(* Logix 5000 project; controller _1407974_PSG_7315 vendor 1 type 14 code 154 rev 20.11; software revision 20.06; part 3 of 4 *)
(* tags used below, declared in another part *)
   AI_L_2_0_Pure_Steam_Conductivity : Analog_Input;
   AI_L_2_1_FW_Press_Low_Warning : OIT_Set_Point_Entry;
   AI_L_2_1_FW_Pressure : Analog_Input;
   AI_R_2_0_Pure_Steam_Temperature : Analog_Input;
   AI_R_2_1_Cond_Pure_Steam_Temperature : Analog_Input;
   Alarm_Pure_Steam_High_Temperature : ALIAS FOR Alarms_Warnings.Latch_Bit[0].4;
   Alarm_Pure_Steam_Temp_Error_Timer : TIMER;
   Alarm_Pure_Steam_Temp_Input_Error : ALIAS FOR Alarms_Warnings.Latch_Bit[0].5;
   Alarm_Pure_Steam_Temp_Input_Error_Ack : ALIAS FOR Alarms_Warnings.Ack[0].5;
   Alarm_Separator_High_Level : ALIAS FOR Alarms_Warnings.Latch_Bit[0].2;
   Alarm_Separator_Low_Level : ALIAS FOR Alarms_Warnings.Latch_Bit[0].3;
   Alarms_Warnings : AW;
   AO_L_3_0_VFD_SPEED : Analog_Output;
   AO_L_3_1_Available : Analog_Output;
   AO_L_3_2_Available : Analog_Output;
   AO_L_3_3_Available : Analog_Output;
   AO_R_4_0_Pure_Steam_Temperature : Analog_Output;
   AO_R_4_1_Available : Analog_Output;
   Cond_Pure_Steam_Hi_Cond_Set_Point_Entry : OIT_Set_Point_Entry;
   Cond_Pure_Steam_Hi_Temp_Set_Point_Entry : OIT_Set_Point_Entry;
   DI_R_1_0_Hi_Hi_Level_LSHH_1950 : ALIAS FOR DI_Remote_1.0;
   DI_R_1_3_Low_Level_LSL_1950 : ALIAS FOR DI_Remote_1.3;
   DI_R_1_4_Air_Low_Pressure_PSL_4030 : ALIAS FOR DI_Remote_1.4;
   DO_L_1_14_Feed_Water_Pump_Contactor : Discrete_Out;
   DO_L_1_1_Alarm_Horn : Discrete_Out;
   DO_L_1_2_Alarm_Light : Discrete_Out;
   DO_Local_1 : INT;
   Feed_Water_Pressure_Set_Point_Entry : OIT_Set_Point_Entry;
   Feedwater_Pressure_PID : PID;
   Free_Run_Pulse_Timer : TIMER;
   FW_Press_PID_Gain_Set_Point_Entry : OIT_Set_Point_Entry;
   FW_Press_PID_Manual_Output_Entry : OIT_Set_Point_Entry;
   FW_Press_PID_Rate_Set_Point_Entry : OIT_Set_Point_Entry;
   FW_Press_PID_Reset_SetPoint_Entry : OIT_Set_Point_Entry;
   FW_Press_PID_Temp_Set_Point_Entry : OIT_Set_Point_Entry;
   Lamp_Test : Push_Button;
   Local_Remote : Latched_Push_Button;
   Low_Feedwater_Pressure : BOOL;
   Network_Ack_All : BOOL;
   Network_Silence : BOOL;
   OIT : OIT_Connections;
   OIT_Auto_Time_Date_Sync : TIMER;
   OIT_Auto_Time_Date_Sync_Interval : TIMER;
   OIT_Day_Set : Push_Button;
   OIT_Hour_Set : Push_Button;
   OIT_Message : OIT_Message;
   OIT_Minute_Set : Push_Button;
   OIT_Month_Set : Push_Button;
   OIT_Year_Set : Push_Button;
   PID_Ramp_Time_Seconds : DINT;
   PID_Ramp_Timer : TIMER;
   Pulse_Bit : BOOL;
   Pure_Steam_High_Temp_Set_Point_Entry : OIT_Set_Point_Entry;
   Pure_Steam_Low_Temp_Set_Point_Entry : OIT_Set_Point_Entry;
   Pure_Steam_Temp_PID_Gain_Set_Point_Entry : OIT_Set_Point_Entry;
   Pure_Steam_Temp_PID_Manual_Output_Entry : OIT_Set_Point_Entry;
   Pure_Steam_Temp_PID_Ramp_Time_Entry : OIT_Set_Point_Entry;
   Pure_Steam_Temp_PID_Rate_Set_Point_Entry : OIT_Set_Point_Entry;
   Pure_Steam_Temp_PID_Reset_SetPoint_Entry : OIT_Set_Point_Entry;
   Pure_Steam_Temp_PID_Temp_Set_Point_Entry : OIT_Set_Point_Entry;
   Pure_Steam_Temperature : PID;
   Pure_Steam_Temperature_Set_Point_Entry : OIT_Set_Point_Entry;
   Read_PLC_Clock : DINT[7];
   Set_PLC_Clock : DINT[7];
   Unit_Hot : BOOL;
   Unit_Status : Unit_Status;
   VFD_Relay_Input : BOOL;
   Warning_Air_Low_Pressure_Timer : TIMER;
   Warning_Cond_Pure_Steam_Analyzer_Fault : ALIAS FOR Alarms_Warnings.Latch_Bit[1].4;
   Warning_Cond_Pure_Steam_Conductivity : ALIAS FOR Alarms_Warnings.Latch_Bit[1].3;
   Warning_Feedwater_Low_Pressure : ALIAS FOR Alarms_Warnings.Latch_Bit[1].9;
   Warning_Feedwater_Press_Low_Pressure_Ack : ALIAS FOR Alarms_Warnings.Ack[1].9;
   Warning_FW_Press_Low_Pressure_Timer : TIMER;
   Warning_Instrument_Air_Low_Pressure : ALIAS FOR Alarms_Warnings.Latch_Bit[1].2;
   Warning_Instrument_Air_Low_Pressure_Ack : ALIAS FOR Alarms_Warnings.Ack[1].2;
   Warning_PLC_OIT_Comm_Counter : COUNTER;
   Warning_PLC_OIT_Comm_Timer : TIMER;
   Warning_PLC_OIT_Commuications_Ack : ALIAS FOR Alarms_Warnings.Ack[1].0;
   Warning_PLC_OIT_Communications : ALIAS FOR Alarms_Warnings.Latch_Bit[1].0;
   Warning_Pure_Steam_Low_Temp_Timer_A : TIMER;
   Warning_Pure_Steam_Low_Temp_Timer_B : TIMER;
   Warning_Pure_Steam_Low_Temperature : ALIAS FOR Alarms_Warnings.Latch_Bit[1].7;
   Warning_Pure_Steam_Low_Temperature_Ack : ALIAS FOR Alarms_Warnings.Ack[1].7;
(* MainProgram, continued *)

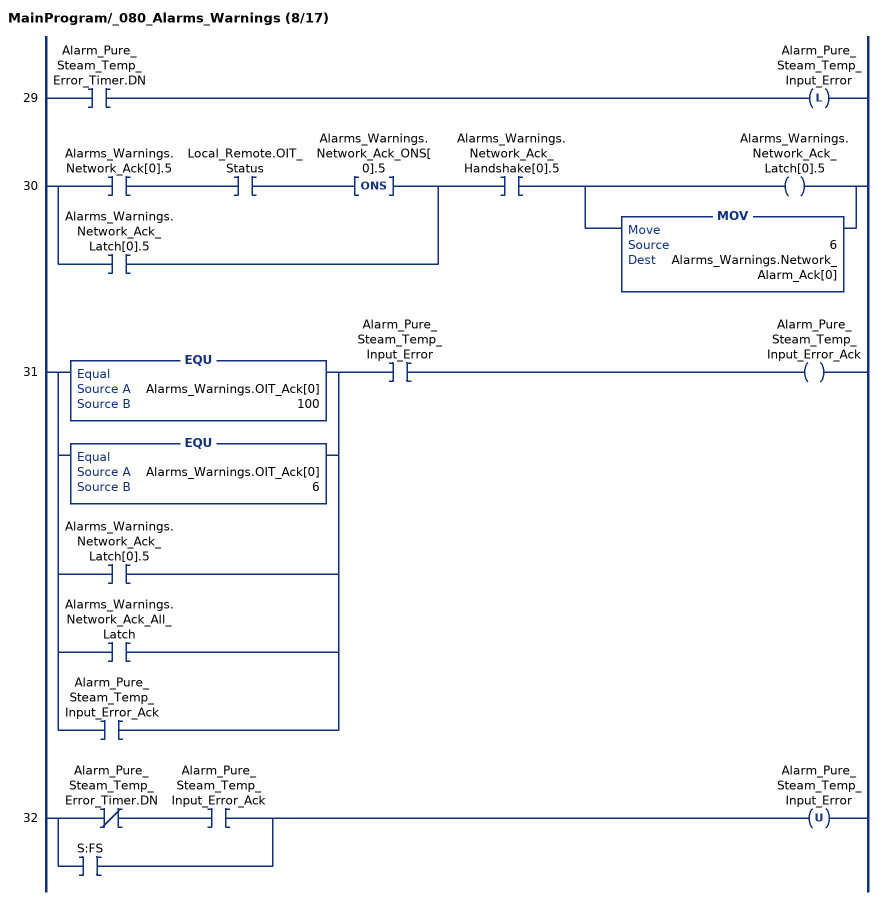
   [picture p43: MainProgram/_080_Alarms_Warnings rungs 29-32]
   29: XIC(Alarm_Pure_Steam_Temp_Error_Timer.DN)OTL(Alarm_Pure_Steam_Temp_Input_Error);
   30: [XIC(Alarms_Warnings.Network_Ack[0].5) XIC(Local_Remote.OIT_Status) ONS(Alarms_Warnings.Network_Ack_ONS[0].5) ,XIC(Alarms_Warnings.Network_Ack_Latch[0].5) ]XIC(Alarms_Warnings.Network_Ack_Handshake[0].5)[OTE(Alarms_Warnings.Network_Ack_Latch[0].5) ,MOV(6,Alarms_Warnings.Network_Alarm_Ack[0]) ];
   31: [EQU(Alarms_Warnings.OIT_Ack[0],100) ,EQU(Alarms_Warnings.OIT_Ack[0],6) ,XIC(Alarms_Warnings.Network_Ack_Latch[0].5) ,XIC(Alarms_Warnings.Network_Ack_All_Latch) ,XIC(Alarm_Pure_Steam_Temp_Input_Error_Ack) ]XIC(Alarm_Pure_Steam_Temp_Input_Error)OTE(Alarm_Pure_Steam_Temp_Input_Error_Ack);
   32: [XIO(Alarm_Pure_Steam_Temp_Error_Timer.DN) XIC(Alarm_Pure_Steam_Temp_Input_Error_Ack) ,XIC(S:FS) ]OTU(Alarm_Pure_Steam_Temp_Input_Error);
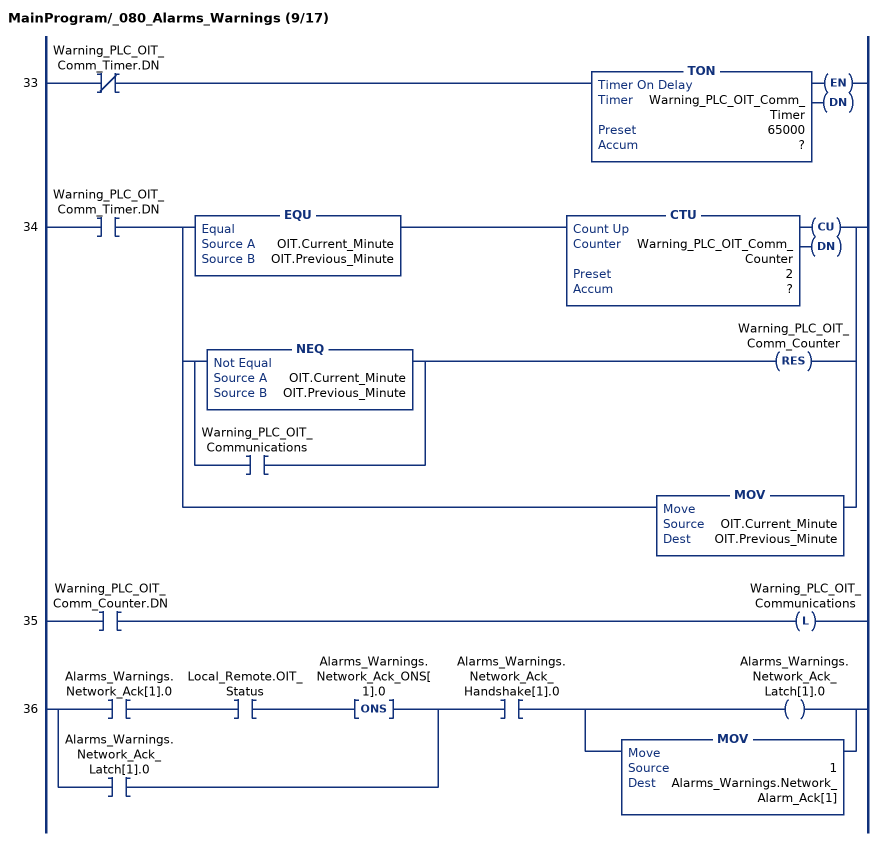
   33: XIO(Warning_PLC_OIT_Comm_Timer.DN)TON(Warning_PLC_OIT_Comm_Timer,?,?);
   34: XIC(Warning_PLC_OIT_Comm_Timer.DN)[EQU(OIT.Current_Minute,OIT.Previous_Minute) CTU(Warning_PLC_OIT_Comm_Counter,?,?) ,[NEQ(OIT.Current_Minute,OIT.Previous_Minute) ,XIC(Warning_PLC_OIT_Communications) ] RES(Warning_PLC_OIT_Comm_Counter) ,MOV(OIT.Current_Minute,OIT.Previous_Minute) ];
   35: XIC(Warning_PLC_OIT_Comm_Counter.DN)OTL(Warning_PLC_OIT_Communications);
   36: [XIC(Alarms_Warnings.Network_Ack[1].0) XIC(Local_Remote.OIT_Status) ONS(Alarms_Warnings.Network_Ack_ONS[1].0) ,XIC(Alarms_Warnings.Network_Ack_Latch[1].0) ]XIC(Alarms_Warnings.Network_Ack_Handshake[1].0)[OTE(Alarms_Warnings.Network_Ack_Latch[1].0) ,MOV(1,Alarms_Warnings.Network_Alarm_Ack[1]) ];
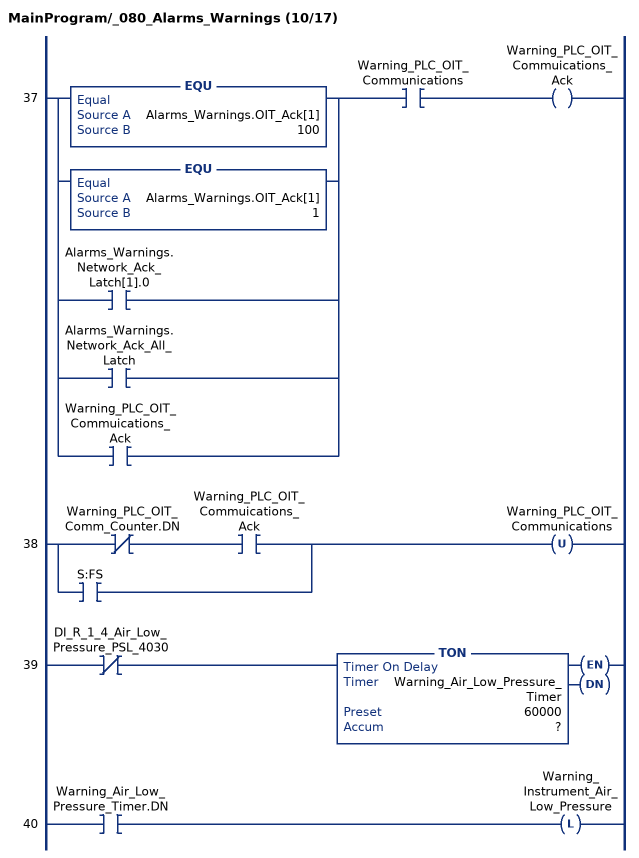
   37: [EQU(Alarms_Warnings.OIT_Ack[1],100) ,EQU(Alarms_Warnings.OIT_Ack[1],1) ,XIC(Alarms_Warnings.Network_Ack_Latch[1].0) ,XIC(Alarms_Warnings.Network_Ack_All_Latch) ,XIC(Warning_PLC_OIT_Commuications_Ack) ]XIC(Warning_PLC_OIT_Communications)OTE(Warning_PLC_OIT_Commuications_Ack);
   38: [XIO(Warning_PLC_OIT_Comm_Counter.DN) XIC(Warning_PLC_OIT_Commuications_Ack) ,XIC(S:FS) ]OTU(Warning_PLC_OIT_Communications);
   39: XIO(DI_R_1_4_Air_Low_Pressure_PSL_4030)TON(Warning_Air_Low_Pressure_Timer,?,?);
   40: XIC(Warning_Air_Low_Pressure_Timer.DN)OTL(Warning_Instrument_Air_Low_Pressure);
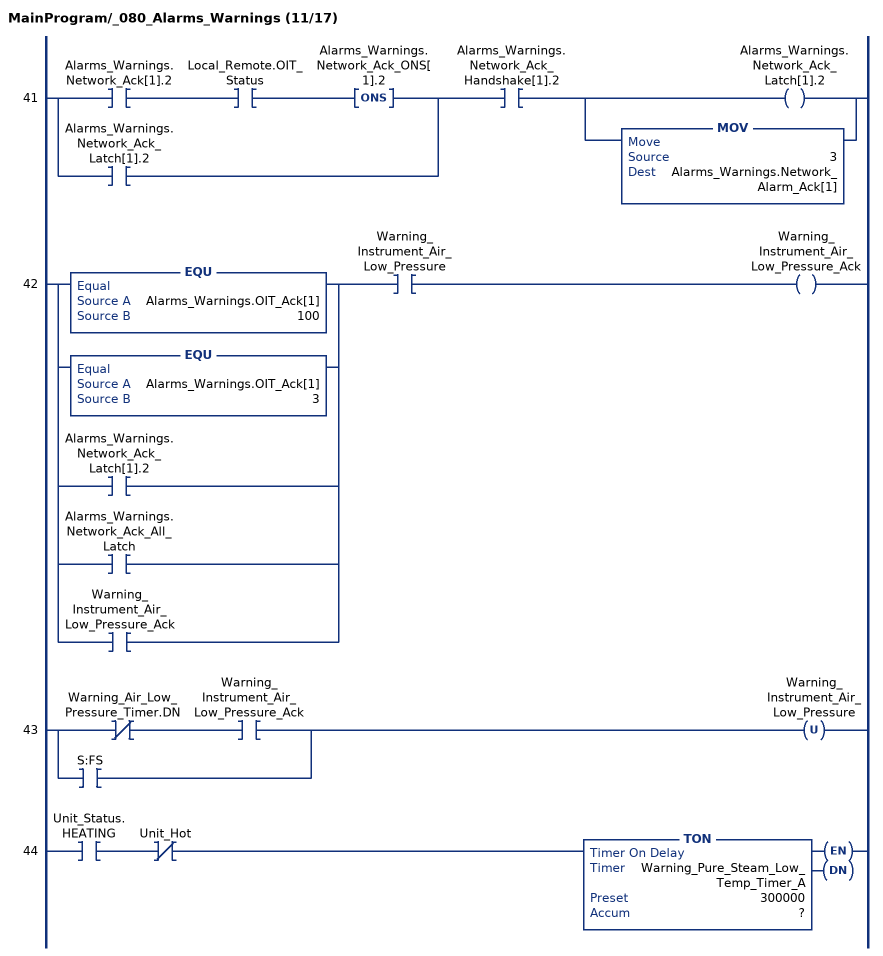
   41: [XIC(Alarms_Warnings.Network_Ack[1].2) XIC(Local_Remote.OIT_Status) ONS(Alarms_Warnings.Network_Ack_ONS[1].2) ,XIC(Alarms_Warnings.Network_Ack_Latch[1].2) ]XIC(Alarms_Warnings.Network_Ack_Handshake[1].2)[OTE(Alarms_Warnings.Network_Ack_Latch[1].2) ,MOV(3,Alarms_Warnings.Network_Alarm_Ack[1]) ];
   42: [EQU(Alarms_Warnings.OIT_Ack[1],100) ,EQU(Alarms_Warnings.OIT_Ack[1],3) ,XIC(Alarms_Warnings.Network_Ack_Latch[1].2) ,XIC(Alarms_Warnings.Network_Ack_All_Latch) ,XIC(Warning_Instrument_Air_Low_Pressure_Ack) ]XIC(Warning_Instrument_Air_Low_Pressure)OTE(Warning_Instrument_Air_Low_Pressure_Ack);
   43: [XIO(Warning_Air_Low_Pressure_Timer.DN) XIC(Warning_Instrument_Air_Low_Pressure_Ack) ,XIC(S:FS) ]OTU(Warning_Instrument_Air_Low_Pressure);
   44: XIC(Unit_Status.HEATING)XIO(Unit_Hot)TON(Warning_Pure_Steam_Low_Temp_Timer_A,?,?);
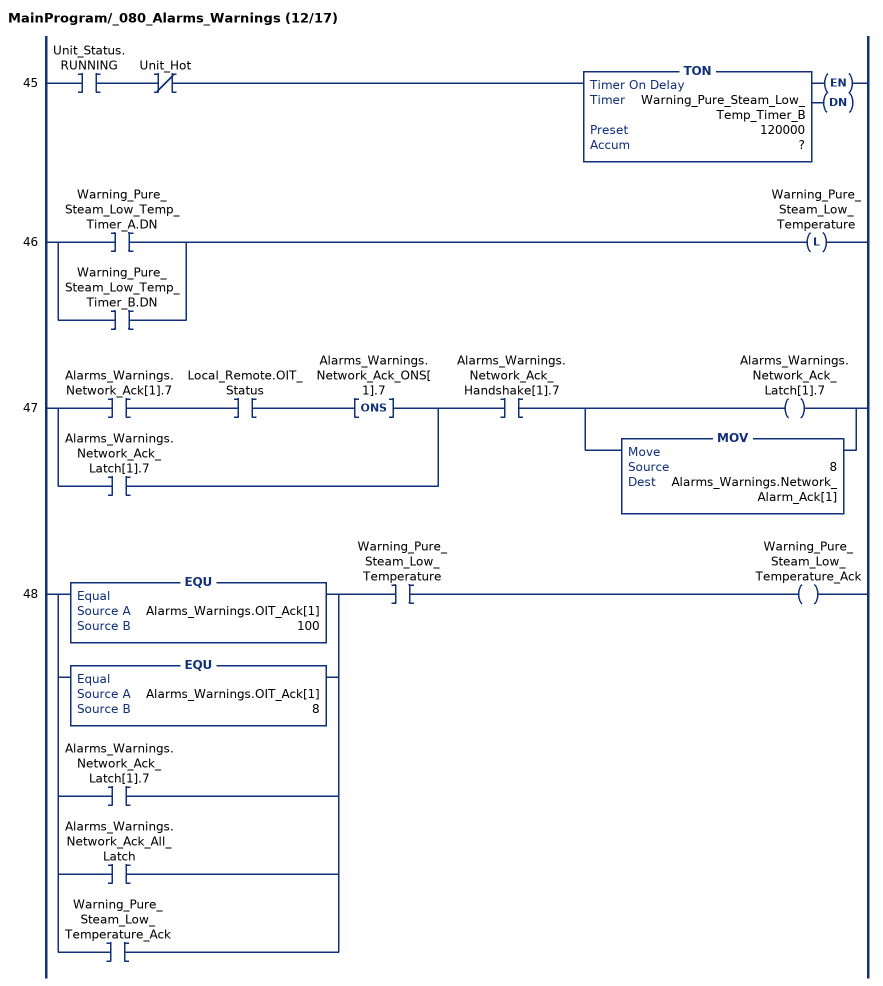
   45: XIC(Unit_Status.RUNNING)XIO(Unit_Hot)TON(Warning_Pure_Steam_Low_Temp_Timer_B,?,?);
   46: [XIC(Warning_Pure_Steam_Low_Temp_Timer_A.DN) ,XIC(Warning_Pure_Steam_Low_Temp_Timer_B.DN) ]OTL(Warning_Pure_Steam_Low_Temperature);
   47: [XIC(Alarms_Warnings.Network_Ack[1].7) XIC(Local_Remote.OIT_Status) ONS(Alarms_Warnings.Network_Ack_ONS[1].7) ,XIC(Alarms_Warnings.Network_Ack_Latch[1].7) ]XIC(Alarms_Warnings.Network_Ack_Handshake[1].7)[OTE(Alarms_Warnings.Network_Ack_Latch[1].7) ,MOV(8,Alarms_Warnings.Network_Alarm_Ack[1]) ];
   48: [EQU(Alarms_Warnings.OIT_Ack[1],100) ,EQU(Alarms_Warnings.OIT_Ack[1],8) ,XIC(Alarms_Warnings.Network_Ack_Latch[1].7) ,XIC(Alarms_Warnings.Network_Ack_All_Latch) ,XIC(Warning_Pure_Steam_Low_Temperature_Ack) ]XIC(Warning_Pure_Steam_Low_Temperature)OTE(Warning_Pure_Steam_Low_Temperature_Ack);
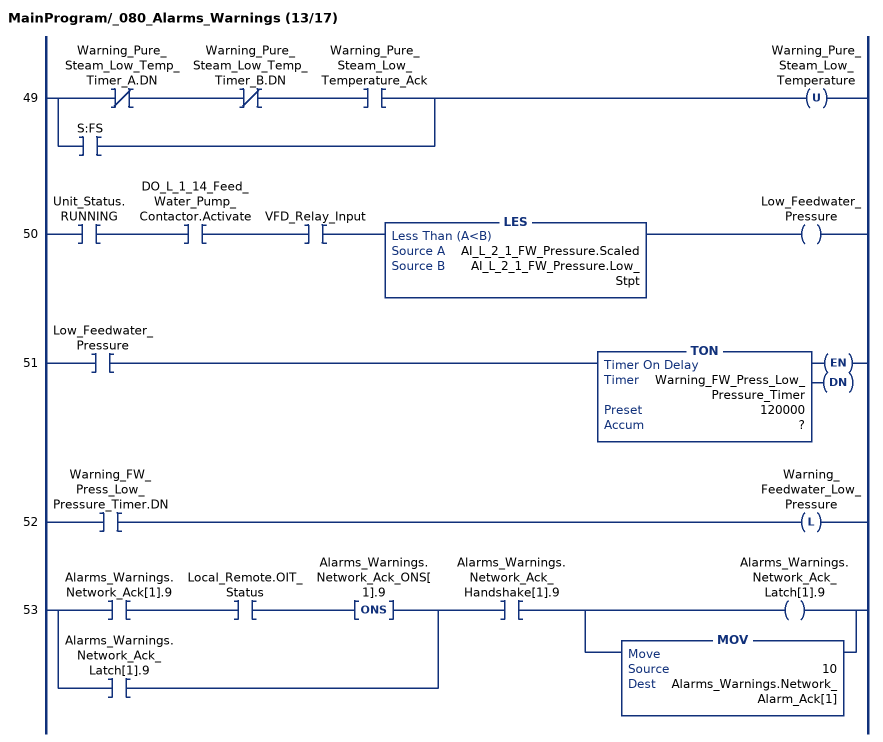
   49: [XIO(Warning_Pure_Steam_Low_Temp_Timer_A.DN) XIO(Warning_Pure_Steam_Low_Temp_Timer_B.DN) XIC(Warning_Pure_Steam_Low_Temperature_Ack) ,XIC(S:FS) ]OTU(Warning_Pure_Steam_Low_Temperature);
   50: XIC(Unit_Status.RUNNING)XIC(DO_L_1_14_Feed_Water_Pump_Contactor.Activate)XIC(VFD_Relay_Input)LES(AI_L_2_1_FW_Pressure.Scaled,AI_L_2_1_FW_Pressure.Low_Stpt)OTE(Low_Feedwater_Pressure);
   51: XIC(Low_Feedwater_Pressure)TON(Warning_FW_Press_Low_Pressure_Timer,?,?);
   52: XIC(Warning_FW_Press_Low_Pressure_Timer.DN)OTL(Warning_Feedwater_Low_Pressure);
   53: [XIC(Alarms_Warnings.Network_Ack[1].9) XIC(Local_Remote.OIT_Status) ONS(Alarms_Warnings.Network_Ack_ONS[1].9) ,XIC(Alarms_Warnings.Network_Ack_Latch[1].9) ]XIC(Alarms_Warnings.Network_Ack_Handshake[1].9)[OTE(Alarms_Warnings.Network_Ack_Latch[1].9) ,MOV(10,Alarms_Warnings.Network_Alarm_Ack[1]) ];
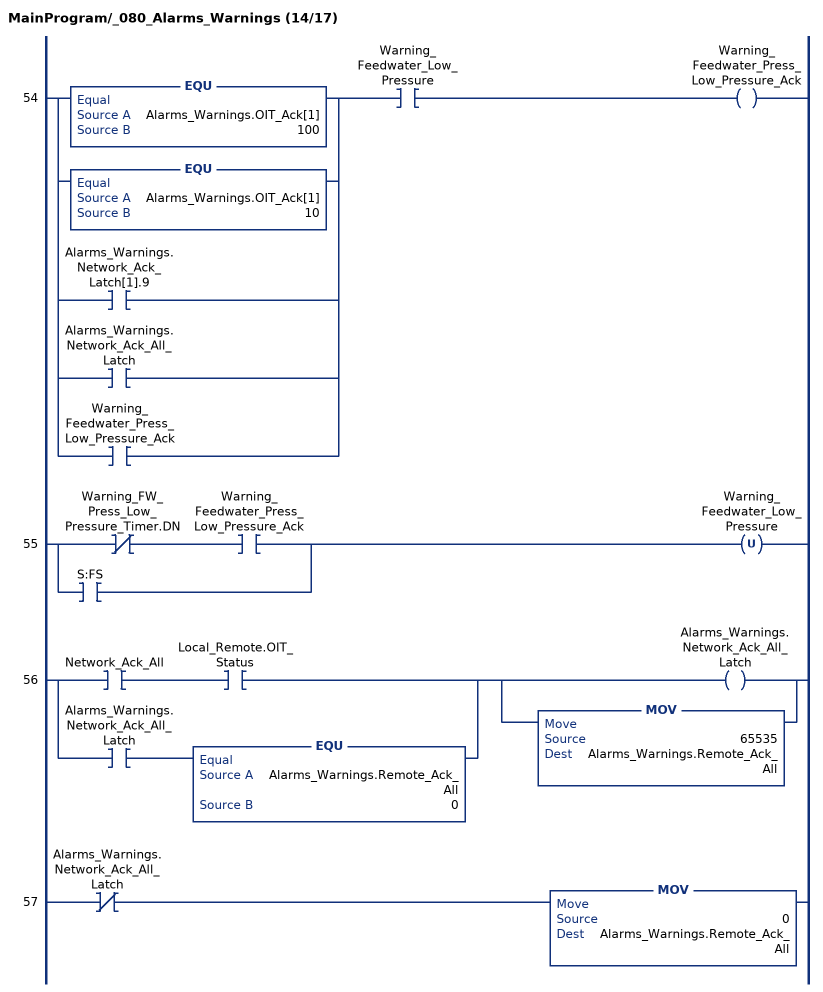
   54: [EQU(Alarms_Warnings.OIT_Ack[1],100) ,EQU(Alarms_Warnings.OIT_Ack[1],10) ,XIC(Alarms_Warnings.Network_Ack_Latch[1].9) ,XIC(Alarms_Warnings.Network_Ack_All_Latch) ,XIC(Warning_Feedwater_Press_Low_Pressure_Ack) ]XIC(Warning_Feedwater_Low_Pressure)OTE(Warning_Feedwater_Press_Low_Pressure_Ack);
   55: [XIO(Warning_FW_Press_Low_Pressure_Timer.DN) XIC(Warning_Feedwater_Press_Low_Pressure_Ack) ,XIC(S:FS) ]OTU(Warning_Feedwater_Low_Pressure);
   56: [XIC(Network_Ack_All) XIC(Local_Remote.OIT_Status) ,XIC(Alarms_Warnings.Network_Ack_All_Latch) EQU(Alarms_Warnings.Remote_Ack_All,0) ][OTE(Alarms_Warnings.Network_Ack_All_Latch) ,MOV(65535,Alarms_Warnings.Remote_Ack_All) ];
   57: XIO(Alarms_Warnings.Network_Ack_All_Latch)MOV(0,Alarms_Warnings.Remote_Ack_All);
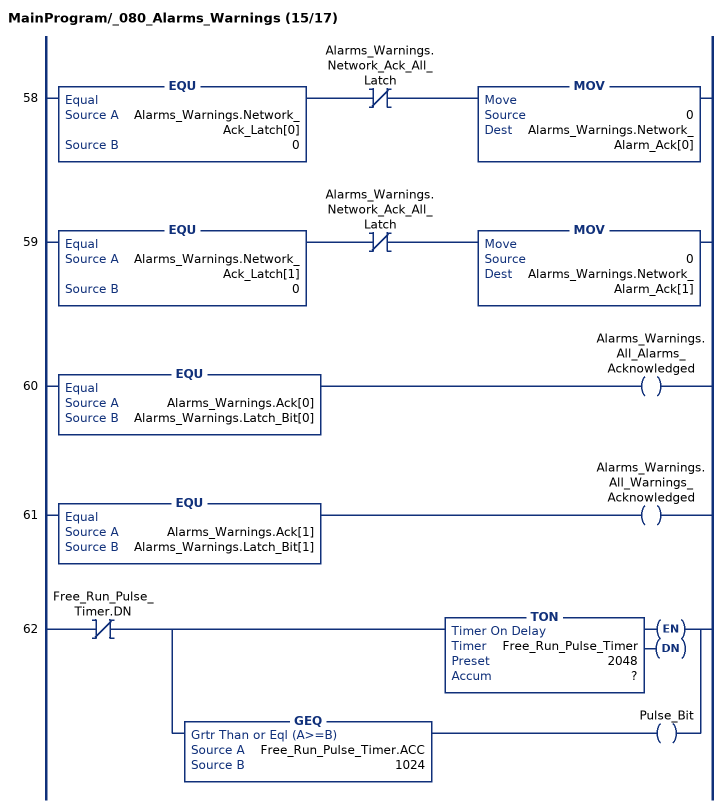
   58: EQU(Alarms_Warnings.Network_Ack_Latch[0],0)XIO(Alarms_Warnings.Network_Ack_All_Latch)MOV(0,Alarms_Warnings.Network_Alarm_Ack[0]);
   59: EQU(Alarms_Warnings.Network_Ack_Latch[1],0)XIO(Alarms_Warnings.Network_Ack_All_Latch)MOV(0,Alarms_Warnings.Network_Alarm_Ack[1]);
   60: EQU(Alarms_Warnings.Ack[0],Alarms_Warnings.Latch_Bit[0])OTE(Alarms_Warnings.All_Alarms_Acknowledged);
   61: EQU(Alarms_Warnings.Ack[1],Alarms_Warnings.Latch_Bit[1])OTE(Alarms_Warnings.All_Warnings_Acknowledged);
   62: XIO(Free_Run_Pulse_Timer.DN)[TON(Free_Run_Pulse_Timer,?,?) ,GEQ(Free_Run_Pulse_Timer.ACC,1024) OTE(Pulse_Bit) ];
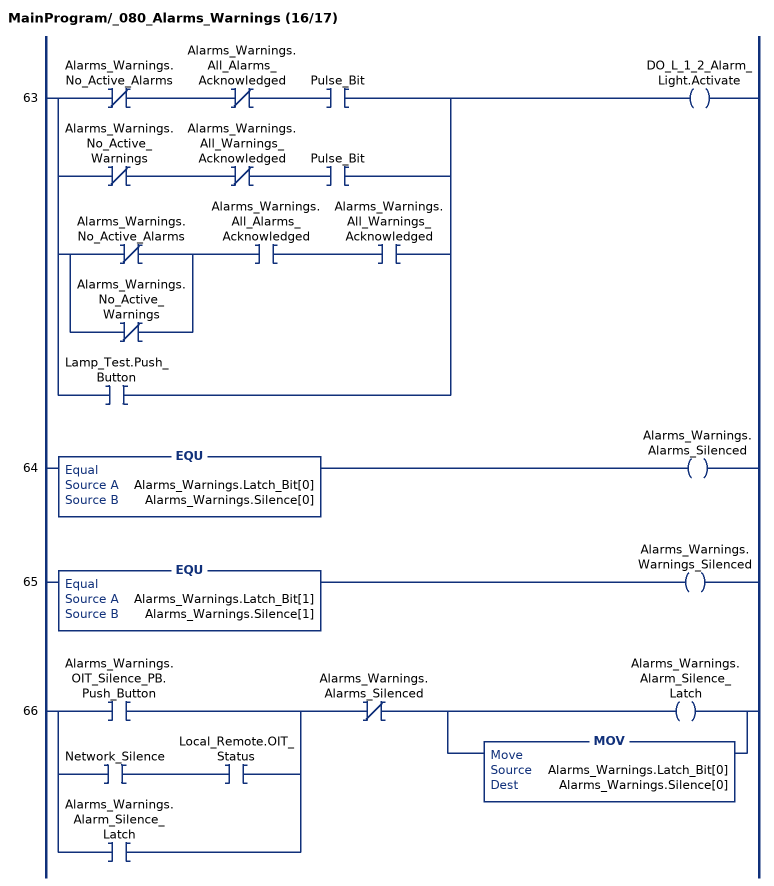
   63: [XIO(Alarms_Warnings.No_Active_Alarms) XIO(Alarms_Warnings.All_Alarms_Acknowledged) XIC(Pulse_Bit) ,XIO(Alarms_Warnings.No_Active_Warnings) XIO(Alarms_Warnings.All_Warnings_Acknowledged) XIC(Pulse_Bit) ,[XIO(Alarms_Warnings.No_Active_Alarms) ,XIO(Alarms_Warnings.No_Active_Warnings) ] XIC(Alarms_Warnings.All_Alarms_Acknowledged) XIC(Alarms_Warnings.All_Warnings_Acknowledged) ,XIC(Lamp_Test.Push_Button) ]OTE(DO_L_1_2_Alarm_Light.Activate);
   64: EQU(Alarms_Warnings.Latch_Bit[0],Alarms_Warnings.Silence[0])OTE(Alarms_Warnings.Alarms_Silenced);
   65: EQU(Alarms_Warnings.Latch_Bit[1],Alarms_Warnings.Silence[1])OTE(Alarms_Warnings.Warnings_Silenced);
   66: [XIC(Alarms_Warnings.OIT_Silence_PB.Push_Button) ,XIC(Network_Silence) XIC(Local_Remote.OIT_Status) ,XIC(Alarms_Warnings.Alarm_Silence_Latch) ]XIO(Alarms_Warnings.Alarms_Silenced)[OTE(Alarms_Warnings.Alarm_Silence_Latch) ,MOV(Alarms_Warnings.Latch_Bit[0],Alarms_Warnings.Silence[0]) ];
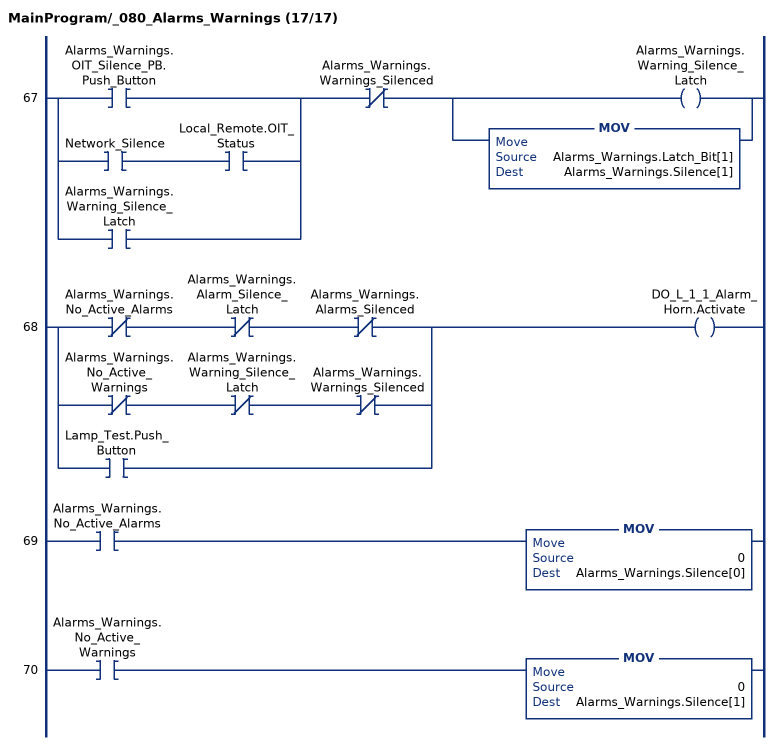
   67: [XIC(Alarms_Warnings.OIT_Silence_PB.Push_Button) ,XIC(Network_Silence) XIC(Local_Remote.OIT_Status) ,XIC(Alarms_Warnings.Warning_Silence_Latch) ]XIO(Alarms_Warnings.Warnings_Silenced)[OTE(Alarms_Warnings.Warning_Silence_Latch) ,MOV(Alarms_Warnings.Latch_Bit[1],Alarms_Warnings.Silence[1]) ];
   68: [XIO(Alarms_Warnings.No_Active_Alarms) XIO(Alarms_Warnings.Alarm_Silence_Latch) XIO(Alarms_Warnings.Alarms_Silenced) ,XIO(Alarms_Warnings.No_Active_Warnings) XIO(Alarms_Warnings.Warning_Silence_Latch) XIO(Alarms_Warnings.Warnings_Silenced) ,XIC(Lamp_Test.Push_Button) ]OTE(DO_L_1_1_Alarm_Horn.Activate);
   69: XIC(Alarms_Warnings.No_Active_Alarms)MOV(0,Alarms_Warnings.Silence[0]);
   70: XIC(Alarms_Warnings.No_Active_Warnings)MOV(0,Alarms_Warnings.Silence[1]);
END_ROUTINE

ROUTINE _090_OIT_Functions   (* ladder *)
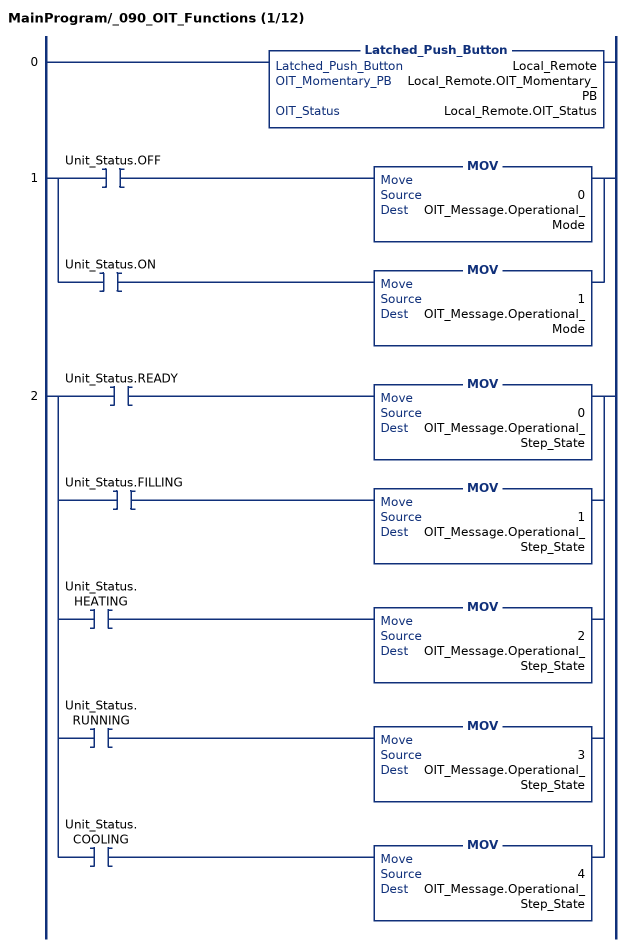
   0: Latched_Push_Button(Local_Remote,Local_Remote.OIT_Momentary_PB,Local_Remote.OIT_Status);
   1: [XIC(Unit_Status.OFF) MOV(0,OIT_Message.Operational_Mode) ,XIC(Unit_Status.ON) MOV(1,OIT_Message.Operational_Mode) ];
   2: [XIC(Unit_Status.READY) MOV(0,OIT_Message.Operational_Step_State) ,XIC(Unit_Status.FILLING) MOV(1,OIT_Message.Operational_Step_State) ,XIC(Unit_Status.HEATING) MOV(2,OIT_Message.Operational_Step_State) ,XIC(Unit_Status.RUNNING) MOV(3,OIT_Message.Operational_Step_State) ,XIC(Unit_Status.COOLING) MOV(4,OIT_Message.Operational_Step_State) ];
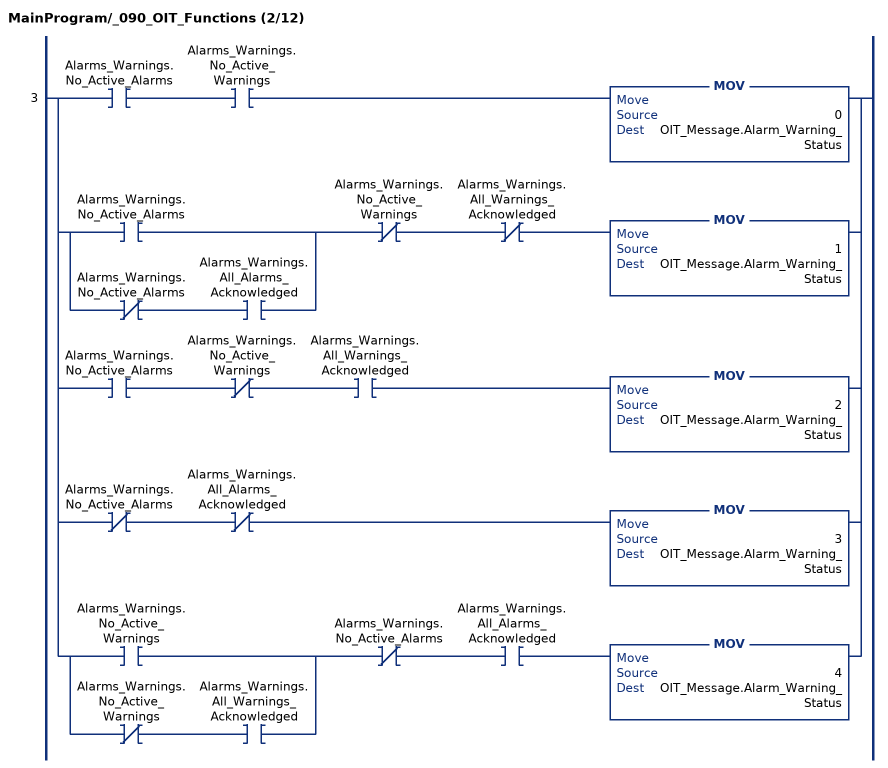
   3: [XIC(Alarms_Warnings.No_Active_Alarms) XIC(Alarms_Warnings.No_Active_Warnings) MOV(0,OIT_Message.Alarm_Warning_Status) ,[XIC(Alarms_Warnings.No_Active_Alarms) ,XIO(Alarms_Warnings.No_Active_Alarms) XIC(Alarms_Warnings.All_Alarms_Acknowledged) ] XIO(Alarms_Warnings.No_Active_Warnings) XIO(Alarms_Warnings.All_Warnings_Acknowledged) MOV(1,OIT_Message.Alarm_Warning_Status) ,XIC(Alarms_Warnings.No_Active_Alarms) XIO(Alarms_Warnings.No_Active_Warnings) XIC(Alarms_Warnings.All_Warnings_Acknowledged) MOV(2,OIT_Message.Alarm_Warning_Status) ,XIO(Alarms_Warnings.No_Active_Alarms) XIO(Alarms_Warnings.All_Alarms_Acknowledged) MOV(3,OIT_Message.Alarm_Warning_Status) ,[XIC(Alarms_Warnings.No_Active_Warnings) ,XIO(Alarms_Warnings.No_Active_Warnings) XIC(Alarms_Warnings.All_Warnings_Acknowledged) ] XIO(Alarms_Warnings.No_Active_Alarms) XIC(Alarms_Warnings.All_Alarms_Acknowledged) MOV(4,OIT_Message.Alarm_Warning_Status) ];
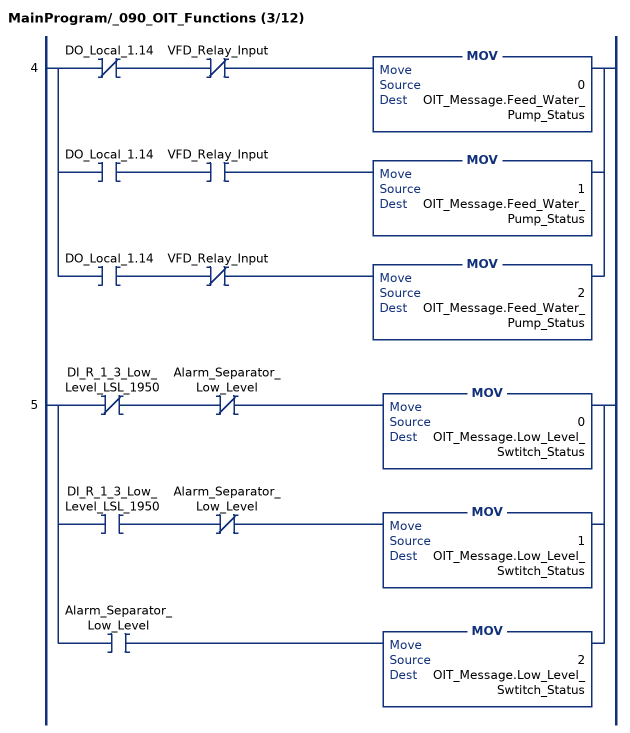
   4: [XIO(DO_Local_1.14) XIO(VFD_Relay_Input) MOV(0,OIT_Message.Feed_Water_Pump_Status) ,XIC(DO_Local_1.14) XIC(VFD_Relay_Input) MOV(1,OIT_Message.Feed_Water_Pump_Status) ,XIC(DO_Local_1.14) XIO(VFD_Relay_Input) MOV(2,OIT_Message.Feed_Water_Pump_Status) ];
   5: [XIO(DI_R_1_3_Low_Level_LSL_1950) XIO(Alarm_Separator_Low_Level) MOV(0,OIT_Message.Low_Level_Swtitch_Status) ,XIC(DI_R_1_3_Low_Level_LSL_1950) XIO(Alarm_Separator_Low_Level) MOV(1,OIT_Message.Low_Level_Swtitch_Status) ,XIC(Alarm_Separator_Low_Level) MOV(2,OIT_Message.Low_Level_Swtitch_Status) ];
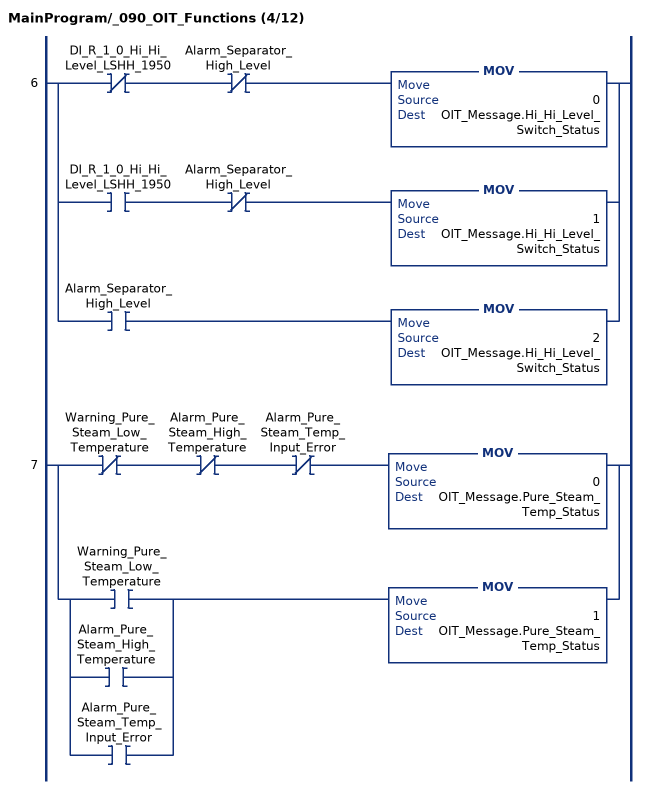
   6: [XIO(DI_R_1_0_Hi_Hi_Level_LSHH_1950) XIO(Alarm_Separator_High_Level) MOV(0,OIT_Message.Hi_Hi_Level_Switch_Status) ,XIC(DI_R_1_0_Hi_Hi_Level_LSHH_1950) XIO(Alarm_Separator_High_Level) MOV(1,OIT_Message.Hi_Hi_Level_Switch_Status) ,XIC(Alarm_Separator_High_Level) MOV(2,OIT_Message.Hi_Hi_Level_Switch_Status) ];
   7: [XIO(Warning_Pure_Steam_Low_Temperature) XIO(Alarm_Pure_Steam_High_Temperature) XIO(Alarm_Pure_Steam_Temp_Input_Error) MOV(0,OIT_Message.Pure_Steam_Temp_Status) ,[XIC(Warning_Pure_Steam_Low_Temperature) ,XIC(Alarm_Pure_Steam_High_Temperature) ,XIC(Alarm_Pure_Steam_Temp_Input_Error) ] MOV(1,OIT_Message.Pure_Steam_Temp_Status) ];
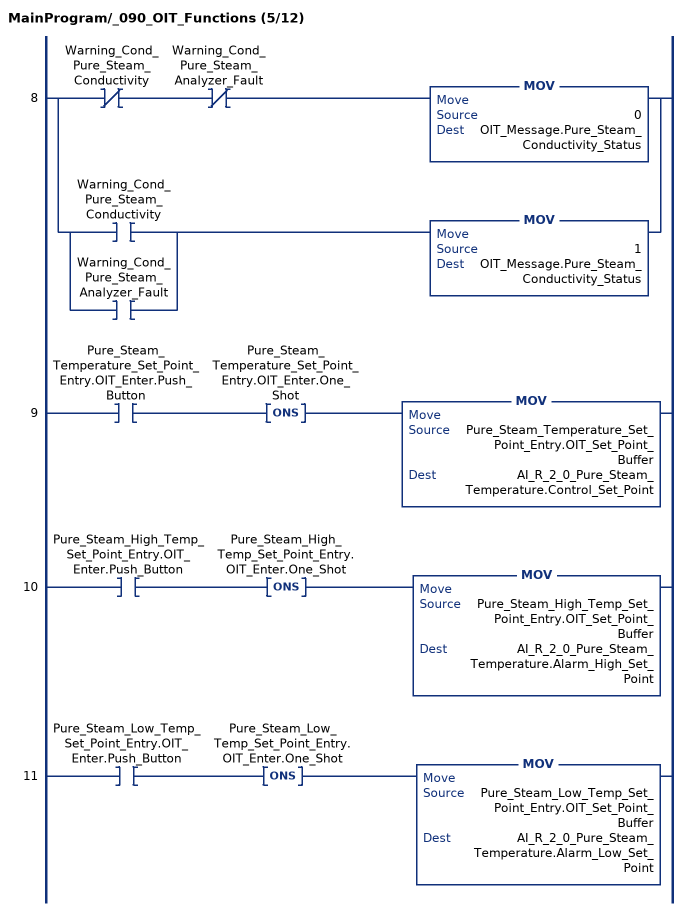
   8: [XIO(Warning_Cond_Pure_Steam_Conductivity) XIO(Warning_Cond_Pure_Steam_Analyzer_Fault) MOV(0,OIT_Message.Pure_Steam_Conductivity_Status) ,[XIC(Warning_Cond_Pure_Steam_Conductivity) ,XIC(Warning_Cond_Pure_Steam_Analyzer_Fault) ] MOV(1,OIT_Message.Pure_Steam_Conductivity_Status) ];
   9: XIC(Pure_Steam_Temperature_Set_Point_Entry.OIT_Enter.Push_Button)ONS(Pure_Steam_Temperature_Set_Point_Entry.OIT_Enter.One_Shot)MOV(Pure_Steam_Temperature_Set_Point_Entry.OIT_Set_Point_Buffer,AI_R_2_0_Pure_Steam_Temperature.Control_Set_Point);
   10: XIC(Pure_Steam_High_Temp_Set_Point_Entry.OIT_Enter.Push_Button)ONS(Pure_Steam_High_Temp_Set_Point_Entry.OIT_Enter.One_Shot)MOV(Pure_Steam_High_Temp_Set_Point_Entry.OIT_Set_Point_Buffer,AI_R_2_0_Pure_Steam_Temperature.Alarm_High_Set_Point);
   11: XIC(Pure_Steam_Low_Temp_Set_Point_Entry.OIT_Enter.Push_Button)ONS(Pure_Steam_Low_Temp_Set_Point_Entry.OIT_Enter.One_Shot)MOV(Pure_Steam_Low_Temp_Set_Point_Entry.OIT_Set_Point_Buffer,AI_R_2_0_Pure_Steam_Temperature.Alarm_Low_Set_Point);
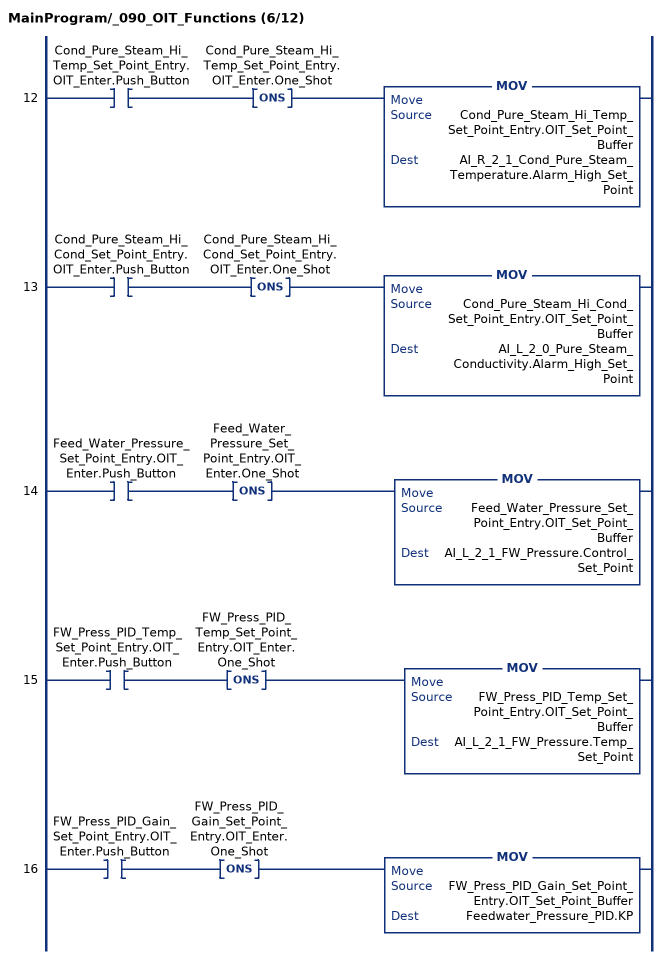
   12: XIC(Cond_Pure_Steam_Hi_Temp_Set_Point_Entry.OIT_Enter.Push_Button)ONS(Cond_Pure_Steam_Hi_Temp_Set_Point_Entry.OIT_Enter.One_Shot)MOV(Cond_Pure_Steam_Hi_Temp_Set_Point_Entry.OIT_Set_Point_Buffer,AI_R_2_1_Cond_Pure_Steam_Temperature.Alarm_High_Set_Point);
   13: XIC(Cond_Pure_Steam_Hi_Cond_Set_Point_Entry.OIT_Enter.Push_Button)ONS(Cond_Pure_Steam_Hi_Cond_Set_Point_Entry.OIT_Enter.One_Shot)MOV(Cond_Pure_Steam_Hi_Cond_Set_Point_Entry.OIT_Set_Point_Buffer,AI_L_2_0_Pure_Steam_Conductivity.Alarm_High_Set_Point);
   14: XIC(Feed_Water_Pressure_Set_Point_Entry.OIT_Enter.Push_Button)ONS(Feed_Water_Pressure_Set_Point_Entry.OIT_Enter.One_Shot)MOV(Feed_Water_Pressure_Set_Point_Entry.OIT_Set_Point_Buffer,AI_L_2_1_FW_Pressure.Control_Set_Point);
   15: XIC(FW_Press_PID_Temp_Set_Point_Entry.OIT_Enter.Push_Button)ONS(FW_Press_PID_Temp_Set_Point_Entry.OIT_Enter.One_Shot)MOV(FW_Press_PID_Temp_Set_Point_Entry.OIT_Set_Point_Buffer,AI_L_2_1_FW_Pressure.Temp_Set_Point);
   16: XIC(FW_Press_PID_Gain_Set_Point_Entry.OIT_Enter.Push_Button)ONS(FW_Press_PID_Gain_Set_Point_Entry.OIT_Enter.One_Shot)MOV(FW_Press_PID_Gain_Set_Point_Entry.OIT_Set_Point_Buffer,Feedwater_Pressure_PID.KP);
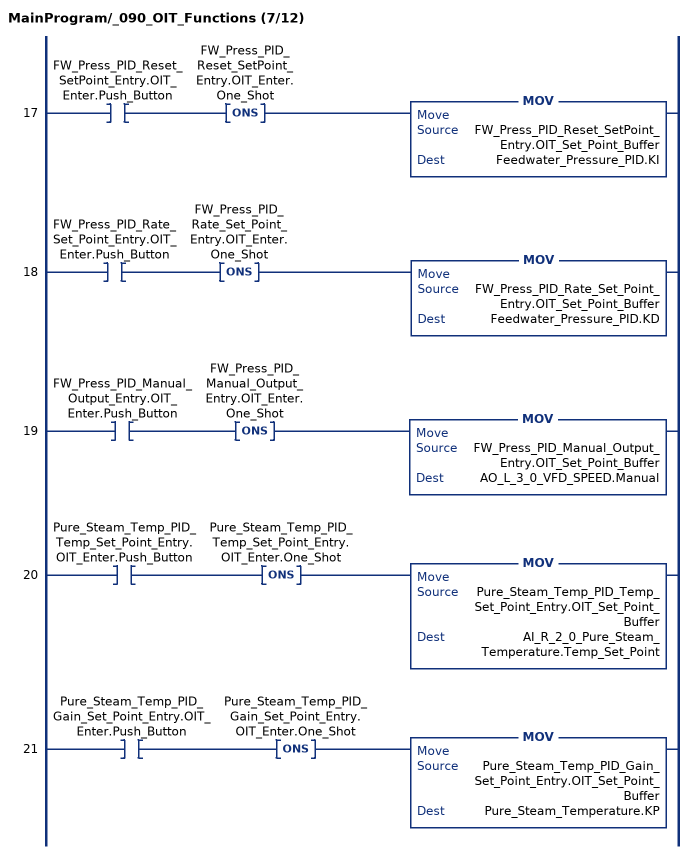
   17: XIC(FW_Press_PID_Reset_SetPoint_Entry.OIT_Enter.Push_Button)ONS(FW_Press_PID_Reset_SetPoint_Entry.OIT_Enter.One_Shot)MOV(FW_Press_PID_Reset_SetPoint_Entry.OIT_Set_Point_Buffer,Feedwater_Pressure_PID.KI);
   18: XIC(FW_Press_PID_Rate_Set_Point_Entry.OIT_Enter.Push_Button)ONS(FW_Press_PID_Rate_Set_Point_Entry.OIT_Enter.One_Shot)MOV(FW_Press_PID_Rate_Set_Point_Entry.OIT_Set_Point_Buffer,Feedwater_Pressure_PID.KD);
   19: XIC(FW_Press_PID_Manual_Output_Entry.OIT_Enter.Push_Button)ONS(FW_Press_PID_Manual_Output_Entry.OIT_Enter.One_Shot)MOV(FW_Press_PID_Manual_Output_Entry.OIT_Set_Point_Buffer,AO_L_3_0_VFD_SPEED.Manual);
   20: XIC(Pure_Steam_Temp_PID_Temp_Set_Point_Entry.OIT_Enter.Push_Button)ONS(Pure_Steam_Temp_PID_Temp_Set_Point_Entry.OIT_Enter.One_Shot)MOV(Pure_Steam_Temp_PID_Temp_Set_Point_Entry.OIT_Set_Point_Buffer,AI_R_2_0_Pure_Steam_Temperature.Temp_Set_Point);
   21: XIC(Pure_Steam_Temp_PID_Gain_Set_Point_Entry.OIT_Enter.Push_Button)ONS(Pure_Steam_Temp_PID_Gain_Set_Point_Entry.OIT_Enter.One_Shot)MOV(Pure_Steam_Temp_PID_Gain_Set_Point_Entry.OIT_Set_Point_Buffer,Pure_Steam_Temperature.KP);
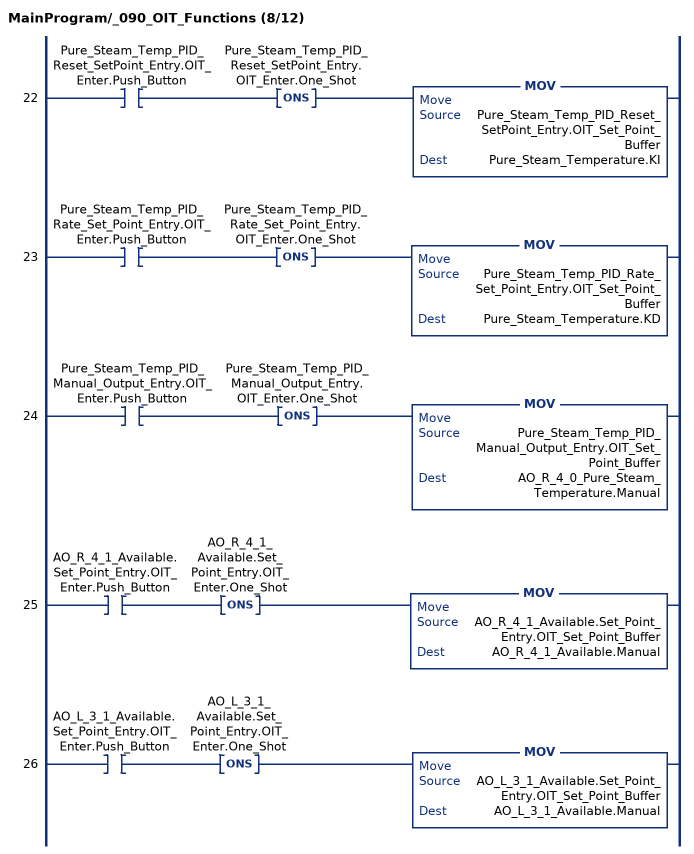
   22: XIC(Pure_Steam_Temp_PID_Reset_SetPoint_Entry.OIT_Enter.Push_Button)ONS(Pure_Steam_Temp_PID_Reset_SetPoint_Entry.OIT_Enter.One_Shot)MOV(Pure_Steam_Temp_PID_Reset_SetPoint_Entry.OIT_Set_Point_Buffer,Pure_Steam_Temperature.KI);
   23: XIC(Pure_Steam_Temp_PID_Rate_Set_Point_Entry.OIT_Enter.Push_Button)ONS(Pure_Steam_Temp_PID_Rate_Set_Point_Entry.OIT_Enter.One_Shot)MOV(Pure_Steam_Temp_PID_Rate_Set_Point_Entry.OIT_Set_Point_Buffer,Pure_Steam_Temperature.KD);
   24: XIC(Pure_Steam_Temp_PID_Manual_Output_Entry.OIT_Enter.Push_Button)ONS(Pure_Steam_Temp_PID_Manual_Output_Entry.OIT_Enter.One_Shot)MOV(Pure_Steam_Temp_PID_Manual_Output_Entry.OIT_Set_Point_Buffer,AO_R_4_0_Pure_Steam_Temperature.Manual);
   25: XIC(AO_R_4_1_Available.Set_Point_Entry.OIT_Enter.Push_Button)ONS(AO_R_4_1_Available.Set_Point_Entry.OIT_Enter.One_Shot)MOV(AO_R_4_1_Available.Set_Point_Entry.OIT_Set_Point_Buffer,AO_R_4_1_Available.Manual);
   26: XIC(AO_L_3_1_Available.Set_Point_Entry.OIT_Enter.Push_Button)ONS(AO_L_3_1_Available.Set_Point_Entry.OIT_Enter.One_Shot)MOV(AO_L_3_1_Available.Set_Point_Entry.OIT_Set_Point_Buffer,AO_L_3_1_Available.Manual);
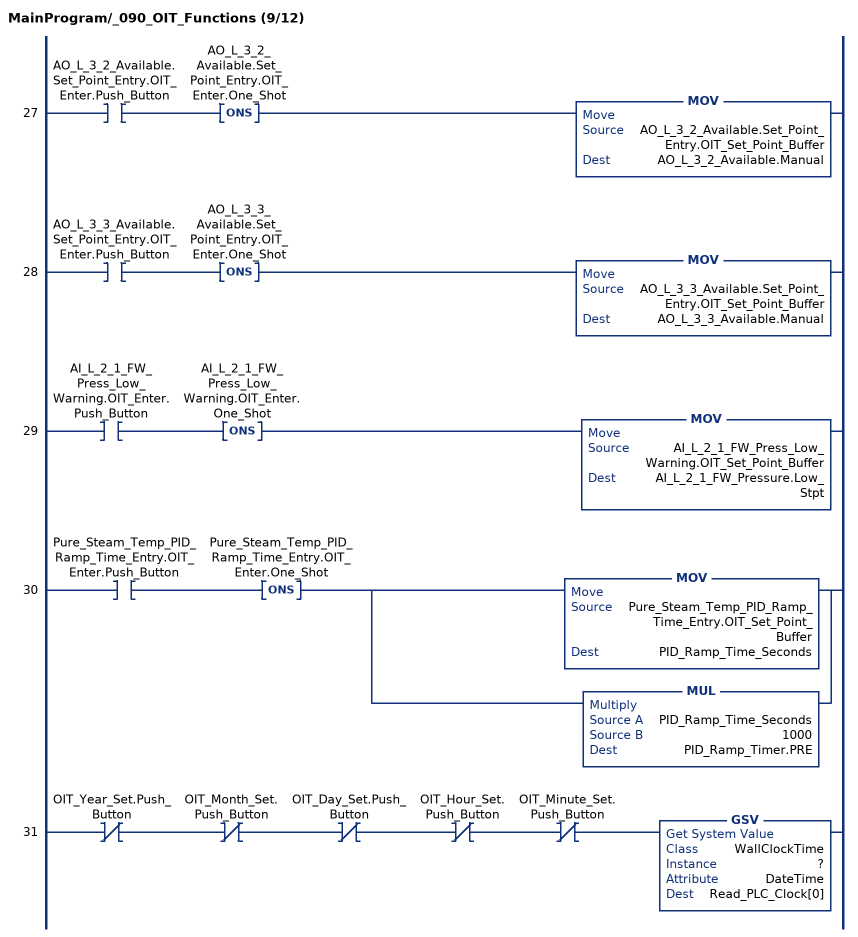
   27: XIC(AO_L_3_2_Available.Set_Point_Entry.OIT_Enter.Push_Button)ONS(AO_L_3_2_Available.Set_Point_Entry.OIT_Enter.One_Shot)MOV(AO_L_3_2_Available.Set_Point_Entry.OIT_Set_Point_Buffer,AO_L_3_2_Available.Manual);
   28: XIC(AO_L_3_3_Available.Set_Point_Entry.OIT_Enter.Push_Button)ONS(AO_L_3_3_Available.Set_Point_Entry.OIT_Enter.One_Shot)MOV(AO_L_3_3_Available.Set_Point_Entry.OIT_Set_Point_Buffer,AO_L_3_3_Available.Manual);
   29: XIC(AI_L_2_1_FW_Press_Low_Warning.OIT_Enter.Push_Button)ONS(AI_L_2_1_FW_Press_Low_Warning.OIT_Enter.One_Shot)MOV(AI_L_2_1_FW_Press_Low_Warning.OIT_Set_Point_Buffer,AI_L_2_1_FW_Pressure.Low_Stpt);
   30: XIC(Pure_Steam_Temp_PID_Ramp_Time_Entry.OIT_Enter.Push_Button)ONS(Pure_Steam_Temp_PID_Ramp_Time_Entry.OIT_Enter.One_Shot)[MOV(Pure_Steam_Temp_PID_Ramp_Time_Entry.OIT_Set_Point_Buffer,PID_Ramp_Time_Seconds) ,MUL(PID_Ramp_Time_Seconds,1000,PID_Ramp_Timer.PRE) ];
   31: XIO(OIT_Year_Set.Push_Button)XIO(OIT_Month_Set.Push_Button)XIO(OIT_Day_Set.Push_Button)XIO(OIT_Hour_Set.Push_Button)XIO(OIT_Minute_Set.Push_Button)GSV(WallClockTime,?,DateTime,Read_PLC_Clock[0]);
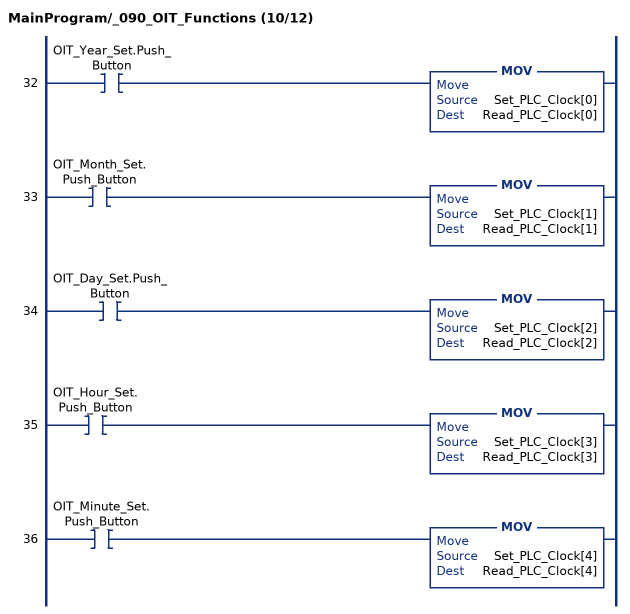
   32: XIC(OIT_Year_Set.Push_Button)MOV(Set_PLC_Clock[0],Read_PLC_Clock[0]);
   33: XIC(OIT_Month_Set.Push_Button)MOV(Set_PLC_Clock[1],Read_PLC_Clock[1]);
   34: XIC(OIT_Day_Set.Push_Button)MOV(Set_PLC_Clock[2],Read_PLC_Clock[2]);
   35: XIC(OIT_Hour_Set.Push_Button)MOV(Set_PLC_Clock[3],Read_PLC_Clock[3]);
   36: XIC(OIT_Minute_Set.Push_Button)MOV(Set_PLC_Clock[4],Read_PLC_Clock[4]);
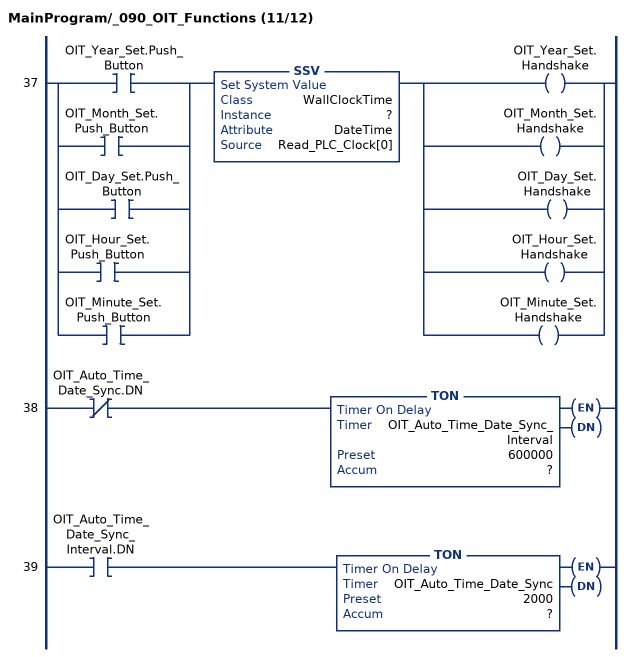
   37: [XIC(OIT_Year_Set.Push_Button) ,XIC(OIT_Month_Set.Push_Button) ,XIC(OIT_Day_Set.Push_Button) ,XIC(OIT_Hour_Set.Push_Button) ,XIC(OIT_Minute_Set.Push_Button) ]SSV(WallClockTime,?,DateTime,Read_PLC_Clock[0])[OTE(OIT_Year_Set.Handshake) ,OTE(OIT_Month_Set.Handshake) ,OTE(OIT_Day_Set.Handshake) ,OTE(OIT_Hour_Set.Handshake) ,OTE(OIT_Minute_Set.Handshake) ];
   38: XIO(OIT_Auto_Time_Date_Sync.DN)TON(OIT_Auto_Time_Date_Sync_Interval,?,?);
   39: XIC(OIT_Auto_Time_Date_Sync_Interval.DN)TON(OIT_Auto_Time_Date_Sync,?,?);
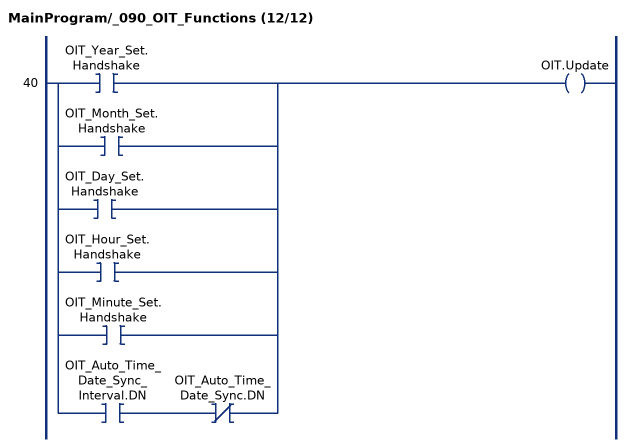
   40: [XIC(OIT_Year_Set.Handshake) ,XIC(OIT_Month_Set.Handshake) ,XIC(OIT_Day_Set.Handshake) ,XIC(OIT_Hour_Set.Handshake) ,XIC(OIT_Minute_Set.Handshake) ,XIC(OIT_Auto_Time_Date_Sync_Interval.DN) XIO(OIT_Auto_Time_Date_Sync.DN) ]OTE(OIT.Update);
END_ROUTINE
